(* IEC 61131-3 sources: STAR-PLC-Agent/results/raw/four_group_20261114/star_deepseek_v4/PUB020/generation/sim_00, 1 file *)

(* ---- test_program.st ---- *)
PROGRAM PLC_PRG
VAR
 BenchStep : UDINT := 0;
 BenchCalls : UDINT := 0;
 BenchDone : BOOL := FALSE;
 BenchUut0 : FB_Task;
 BenchUut1 : FB_Task;
 TraceIn_Mode : ARRAY[0..14] OF BOOL;
 TraceIn_ForwardButton : ARRAY[0..14] OF BOOL;
 TraceIn_ReverseButton : ARRAY[0..14] OF BOOL;
 TraceIn_SensorFeed : ARRAY[0..14] OF BOOL;
 TraceIn_SensorWash : ARRAY[0..14] OF BOOL;
 TraceIn_SensorWeight : ARRAY[0..14] OF BOOL;
 TraceIn_SensorFiring : ARRAY[0..14] OF BOOL;
 TraceIn_SensorOutput : ARRAY[0..14] OF BOOL;
 TraceIn_washComplete : ARRAY[0..14] OF BOOL;
 TraceIn_weightComplete : ARRAY[0..14] OF BOOL;
 TraceIn_weight : ARRAY[0..14] OF REAL;
 TraceIn_firingComplete : ARRAY[0..14] OF BOOL;
 TraceOut_MotorForward : ARRAY[0..14] OF BOOL;
 TraceOut_MotorReverse : ARRAY[0..14] OF BOOL;
 TraceOut_kick : ARRAY[0..14] OF BOOL;
 TraceOut_CompletionLight : ARRAY[0..14] OF BOOL;
 TraceOut_firingTemp : ARRAY[0..14] OF REAL;
END_VAR

IF NOT BenchDone THEN
 CASE BenchStep OF
 0:
   BenchUut0.Mode := TRUE;
   BenchUut0.ForwardButton := FALSE;
   BenchUut0.ReverseButton := FALSE;
   BenchUut0.SensorFeed := TRUE;
   BenchUut0.SensorWash := FALSE;
   BenchUut0.SensorWeight := FALSE;
   BenchUut0.SensorFiring := FALSE;
   BenchUut0.SensorOutput := FALSE;
   BenchUut0.washComplete := FALSE;
   BenchUut0.weightComplete := FALSE;
   BenchUut0.weight := REAL#0.0;
   BenchUut0.firingComplete := FALSE;
   TraceIn_Mode[0] := BenchUut0.Mode;
   TraceIn_ForwardButton[0] := BenchUut0.ForwardButton;
   TraceIn_ReverseButton[0] := BenchUut0.ReverseButton;
   TraceIn_SensorFeed[0] := BenchUut0.SensorFeed;
   TraceIn_SensorWash[0] := BenchUut0.SensorWash;
   TraceIn_SensorWeight[0] := BenchUut0.SensorWeight;
   TraceIn_SensorFiring[0] := BenchUut0.SensorFiring;
   TraceIn_SensorOutput[0] := BenchUut0.SensorOutput;
   TraceIn_washComplete[0] := BenchUut0.washComplete;
   TraceIn_weightComplete[0] := BenchUut0.weightComplete;
   TraceIn_weight[0] := BenchUut0.weight;
   TraceIn_firingComplete[0] := BenchUut0.firingComplete;
   BenchUut0();
   TraceOut_MotorForward[0] := BenchUut0.MotorForward;
   TraceOut_MotorReverse[0] := BenchUut0.MotorReverse;
   TraceOut_kick[0] := BenchUut0.kick;
   TraceOut_CompletionLight[0] := BenchUut0.CompletionLight;
   TraceOut_firingTemp[0] := BenchUut0.firingTemp;
   BenchCalls := BenchCalls + 1;
 1:
   BenchUut0.Mode := TRUE;
   BenchUut0.ForwardButton := FALSE;
   BenchUut0.ReverseButton := FALSE;
   BenchUut0.SensorFeed := FALSE;
   BenchUut0.SensorWash := TRUE;
   BenchUut0.SensorWeight := FALSE;
   BenchUut0.SensorFiring := FALSE;
   BenchUut0.SensorOutput := FALSE;
   BenchUut0.washComplete := FALSE;
   BenchUut0.weightComplete := FALSE;
   BenchUut0.weight := REAL#0.0;
   BenchUut0.firingComplete := FALSE;
   TraceIn_Mode[1] := BenchUut0.Mode;
   TraceIn_ForwardButton[1] := BenchUut0.ForwardButton;
   TraceIn_ReverseButton[1] := BenchUut0.ReverseButton;
   TraceIn_SensorFeed[1] := BenchUut0.SensorFeed;
   TraceIn_SensorWash[1] := BenchUut0.SensorWash;
   TraceIn_SensorWeight[1] := BenchUut0.SensorWeight;
   TraceIn_SensorFiring[1] := BenchUut0.SensorFiring;
   TraceIn_SensorOutput[1] := BenchUut0.SensorOutput;
   TraceIn_washComplete[1] := BenchUut0.washComplete;
   TraceIn_weightComplete[1] := BenchUut0.weightComplete;
   TraceIn_weight[1] := BenchUut0.weight;
   TraceIn_firingComplete[1] := BenchUut0.firingComplete;
   BenchUut0();
   TraceOut_MotorForward[1] := BenchUut0.MotorForward;
   TraceOut_MotorReverse[1] := BenchUut0.MotorReverse;
   TraceOut_kick[1] := BenchUut0.kick;
   TraceOut_CompletionLight[1] := BenchUut0.CompletionLight;
   TraceOut_firingTemp[1] := BenchUut0.firingTemp;
   BenchCalls := BenchCalls + 1;
 2:
   BenchUut0.Mode := TRUE;
   BenchUut0.ForwardButton := FALSE;
   BenchUut0.ReverseButton := FALSE;
   BenchUut0.SensorFeed := FALSE;
   BenchUut0.SensorWash := TRUE;
   BenchUut0.SensorWeight := FALSE;
   BenchUut0.SensorFiring := FALSE;
   BenchUut0.SensorOutput := FALSE;
   BenchUut0.washComplete := TRUE;
   BenchUut0.weightComplete := FALSE;
   BenchUut0.weight := REAL#0.0;
   BenchUut0.firingComplete := FALSE;
   TraceIn_Mode[2] := BenchUut0.Mode;
   TraceIn_ForwardButton[2] := BenchUut0.ForwardButton;
   TraceIn_ReverseButton[2] := BenchUut0.ReverseButton;
   TraceIn_SensorFeed[2] := BenchUut0.SensorFeed;
   TraceIn_SensorWash[2] := BenchUut0.SensorWash;
   TraceIn_SensorWeight[2] := BenchUut0.SensorWeight;
   TraceIn_SensorFiring[2] := BenchUut0.SensorFiring;
   TraceIn_SensorOutput[2] := BenchUut0.SensorOutput;
   TraceIn_washComplete[2] := BenchUut0.washComplete;
   TraceIn_weightComplete[2] := BenchUut0.weightComplete;
   TraceIn_weight[2] := BenchUut0.weight;
   TraceIn_firingComplete[2] := BenchUut0.firingComplete;
   BenchUut0();
   TraceOut_MotorForward[2] := BenchUut0.MotorForward;
   TraceOut_MotorReverse[2] := BenchUut0.MotorReverse;
   TraceOut_kick[2] := BenchUut0.kick;
   TraceOut_CompletionLight[2] := BenchUut0.CompletionLight;
   TraceOut_firingTemp[2] := BenchUut0.firingTemp;
   BenchCalls := BenchCalls + 1;
 3:
   BenchUut0.Mode := TRUE;
   BenchUut0.ForwardButton := FALSE;
   BenchUut0.ReverseButton := FALSE;
   BenchUut0.SensorFeed := FALSE;
   BenchUut0.SensorWash := FALSE;
   BenchUut0.SensorWeight := TRUE;
   BenchUut0.SensorFiring := FALSE;
   BenchUut0.SensorOutput := FALSE;
   BenchUut0.washComplete := FALSE;
   BenchUut0.weightComplete := FALSE;
   BenchUut0.weight := REAL#0.0;
   BenchUut0.firingComplete := FALSE;
   TraceIn_Mode[3] := BenchUut0.Mode;
   TraceIn_ForwardButton[3] := BenchUut0.ForwardButton;
   TraceIn_ReverseButton[3] := BenchUut0.ReverseButton;
   TraceIn_SensorFeed[3] := BenchUut0.SensorFeed;
   TraceIn_SensorWash[3] := BenchUut0.SensorWash;
   TraceIn_SensorWeight[3] := BenchUut0.SensorWeight;
   TraceIn_SensorFiring[3] := BenchUut0.SensorFiring;
   TraceIn_SensorOutput[3] := BenchUut0.SensorOutput;
   TraceIn_washComplete[3] := BenchUut0.washComplete;
   TraceIn_weightComplete[3] := BenchUut0.weightComplete;
   TraceIn_weight[3] := BenchUut0.weight;
   TraceIn_firingComplete[3] := BenchUut0.firingComplete;
   BenchUut0();
   TraceOut_MotorForward[3] := BenchUut0.MotorForward;
   TraceOut_MotorReverse[3] := BenchUut0.MotorReverse;
   TraceOut_kick[3] := BenchUut0.kick;
   TraceOut_CompletionLight[3] := BenchUut0.CompletionLight;
   TraceOut_firingTemp[3] := BenchUut0.firingTemp;
   BenchCalls := BenchCalls + 1;
 4:
   BenchUut0.Mode := TRUE;
   BenchUut0.ForwardButton := FALSE;
   BenchUut0.ReverseButton := FALSE;
   BenchUut0.SensorFeed := FALSE;
   BenchUut0.SensorWash := FALSE;
   BenchUut0.SensorWeight := TRUE;
   BenchUut0.SensorFiring := FALSE;
   BenchUut0.SensorOutput := FALSE;
   BenchUut0.washComplete := FALSE;
   BenchUut0.weightComplete := TRUE;
   BenchUut0.weight := REAL#200.0;
   BenchUut0.firingComplete := FALSE;
   TraceIn_Mode[4] := BenchUut0.Mode;
   TraceIn_ForwardButton[4] := BenchUut0.ForwardButton;
   TraceIn_ReverseButton[4] := BenchUut0.ReverseButton;
   TraceIn_SensorFeed[4] := BenchUut0.SensorFeed;
   TraceIn_SensorWash[4] := BenchUut0.SensorWash;
   TraceIn_SensorWeight[4] := BenchUut0.SensorWeight;
   TraceIn_SensorFiring[4] := BenchUut0.SensorFiring;
   TraceIn_SensorOutput[4] := BenchUut0.SensorOutput;
   TraceIn_washComplete[4] := BenchUut0.washComplete;
   TraceIn_weightComplete[4] := BenchUut0.weightComplete;
   TraceIn_weight[4] := BenchUut0.weight;
   TraceIn_firingComplete[4] := BenchUut0.firingComplete;
   BenchUut0();
   TraceOut_MotorForward[4] := BenchUut0.MotorForward;
   TraceOut_MotorReverse[4] := BenchUut0.MotorReverse;
   TraceOut_kick[4] := BenchUut0.kick;
   TraceOut_CompletionLight[4] := BenchUut0.CompletionLight;
   TraceOut_firingTemp[4] := BenchUut0.firingTemp;
   BenchCalls := BenchCalls + 1;
 5:
   BenchUut0.Mode := TRUE;
   BenchUut0.ForwardButton := FALSE;
   BenchUut0.ReverseButton := FALSE;
   BenchUut0.SensorFeed := FALSE;
   BenchUut0.SensorWash := FALSE;
   BenchUut0.SensorWeight := FALSE;
   BenchUut0.SensorFiring := TRUE;
   BenchUut0.SensorOutput := FALSE;
   BenchUut0.washComplete := FALSE;
   BenchUut0.weightComplete := FALSE;
   BenchUut0.weight := REAL#200.0;
   BenchUut0.firingComplete := FALSE;
   TraceIn_Mode[5] := BenchUut0.Mode;
   TraceIn_ForwardButton[5] := BenchUut0.ForwardButton;
   TraceIn_ReverseButton[5] := BenchUut0.ReverseButton;
   TraceIn_SensorFeed[5] := BenchUut0.SensorFeed;
   TraceIn_SensorWash[5] := BenchUut0.SensorWash;
   TraceIn_SensorWeight[5] := BenchUut0.SensorWeight;
   TraceIn_SensorFiring[5] := BenchUut0.SensorFiring;
   TraceIn_SensorOutput[5] := BenchUut0.SensorOutput;
   TraceIn_washComplete[5] := BenchUut0.washComplete;
   TraceIn_weightComplete[5] := BenchUut0.weightComplete;
   TraceIn_weight[5] := BenchUut0.weight;
   TraceIn_firingComplete[5] := BenchUut0.firingComplete;
   BenchUut0();
   TraceOut_MotorForward[5] := BenchUut0.MotorForward;
   TraceOut_MotorReverse[5] := BenchUut0.MotorReverse;
   TraceOut_kick[5] := BenchUut0.kick;
   TraceOut_CompletionLight[5] := BenchUut0.CompletionLight;
   TraceOut_firingTemp[5] := BenchUut0.firingTemp;
   BenchCalls := BenchCalls + 1;
 6:
   BenchUut0.Mode := TRUE;
   BenchUut0.ForwardButton := FALSE;
   BenchUut0.ReverseButton := FALSE;
   BenchUut0.SensorFeed := FALSE;
   BenchUut0.SensorWash := FALSE;
   BenchUut0.SensorWeight := FALSE;
   BenchUut0.SensorFiring := TRUE;
   BenchUut0.SensorOutput := FALSE;
   BenchUut0.washComplete := FALSE;
   BenchUut0.weightComplete := FALSE;
   BenchUut0.weight := REAL#200.0;
   BenchUut0.firingComplete := TRUE;
   TraceIn_Mode[6] := BenchUut0.Mode;
   TraceIn_ForwardButton[6] := BenchUut0.ForwardButton;
   TraceIn_ReverseButton[6] := BenchUut0.ReverseButton;
   TraceIn_SensorFeed[6] := BenchUut0.SensorFeed;
   TraceIn_SensorWash[6] := BenchUut0.SensorWash;
   TraceIn_SensorWeight[6] := BenchUut0.SensorWeight;
   TraceIn_SensorFiring[6] := BenchUut0.SensorFiring;
   TraceIn_SensorOutput[6] := BenchUut0.SensorOutput;
   TraceIn_washComplete[6] := BenchUut0.washComplete;
   TraceIn_weightComplete[6] := BenchUut0.weightComplete;
   TraceIn_weight[6] := BenchUut0.weight;
   TraceIn_firingComplete[6] := BenchUut0.firingComplete;
   BenchUut0();
   TraceOut_MotorForward[6] := BenchUut0.MotorForward;
   TraceOut_MotorReverse[6] := BenchUut0.MotorReverse;
   TraceOut_kick[6] := BenchUut0.kick;
   TraceOut_CompletionLight[6] := BenchUut0.CompletionLight;
   TraceOut_firingTemp[6] := BenchUut0.firingTemp;
   BenchCalls := BenchCalls + 1;
 7:
   BenchUut0.Mode := TRUE;
   BenchUut0.ForwardButton := FALSE;
   BenchUut0.ReverseButton := FALSE;
   BenchUut0.SensorFeed := FALSE;
   BenchUut0.SensorWash := FALSE;
   BenchUut0.SensorWeight := FALSE;
   BenchUut0.SensorFiring := FALSE;
   BenchUut0.SensorOutput := TRUE;
   BenchUut0.washComplete := FALSE;
   BenchUut0.weightComplete := FALSE;
   BenchUut0.weight := REAL#200.0;
   BenchUut0.firingComplete := FALSE;
   TraceIn_Mode[7] := BenchUut0.Mode;
   TraceIn_ForwardButton[7] := BenchUut0.ForwardButton;
   TraceIn_ReverseButton[7] := BenchUut0.ReverseButton;
   TraceIn_SensorFeed[7] := BenchUut0.SensorFeed;
   TraceIn_SensorWash[7] := BenchUut0.SensorWash;
   TraceIn_SensorWeight[7] := BenchUut0.SensorWeight;
   TraceIn_SensorFiring[7] := BenchUut0.SensorFiring;
   TraceIn_SensorOutput[7] := BenchUut0.SensorOutput;
   TraceIn_washComplete[7] := BenchUut0.washComplete;
   TraceIn_weightComplete[7] := BenchUut0.weightComplete;
   TraceIn_weight[7] := BenchUut0.weight;
   TraceIn_firingComplete[7] := BenchUut0.firingComplete;
   BenchUut0();
   TraceOut_MotorForward[7] := BenchUut0.MotorForward;
   TraceOut_MotorReverse[7] := BenchUut0.MotorReverse;
   TraceOut_kick[7] := BenchUut0.kick;
   TraceOut_CompletionLight[7] := BenchUut0.CompletionLight;
   TraceOut_firingTemp[7] := BenchUut0.firingTemp;
   BenchCalls := BenchCalls + 1;
 8:
   BenchUut1.Mode := TRUE;
   BenchUut1.ForwardButton := FALSE;
   BenchUut1.ReverseButton := FALSE;
   BenchUut1.SensorFeed := TRUE;
   BenchUut1.SensorWash := FALSE;
   BenchUut1.SensorWeight := FALSE;
   BenchUut1.SensorFiring := FALSE;
   BenchUut1.SensorOutput := FALSE;
   BenchUut1.washComplete := FALSE;
   BenchUut1.weightComplete := FALSE;
   BenchUut1.weight := REAL#0.0;
   BenchUut1.firingComplete := FALSE;
   TraceIn_Mode[8] := BenchUut1.Mode;
   TraceIn_ForwardButton[8] := BenchUut1.ForwardButton;
   TraceIn_ReverseButton[8] := BenchUut1.ReverseButton;
   TraceIn_SensorFeed[8] := BenchUut1.SensorFeed;
   TraceIn_SensorWash[8] := BenchUut1.SensorWash;
   TraceIn_SensorWeight[8] := BenchUut1.SensorWeight;
   TraceIn_SensorFiring[8] := BenchUut1.SensorFiring;
   TraceIn_SensorOutput[8] := BenchUut1.SensorOutput;
   TraceIn_washComplete[8] := BenchUut1.washComplete;
   TraceIn_weightComplete[8] := BenchUut1.weightComplete;
   TraceIn_weight[8] := BenchUut1.weight;
   TraceIn_firingComplete[8] := BenchUut1.firingComplete;
   BenchUut1();
   TraceOut_MotorForward[8] := BenchUut1.MotorForward;
   TraceOut_MotorReverse[8] := BenchUut1.MotorReverse;
   TraceOut_kick[8] := BenchUut1.kick;
   TraceOut_CompletionLight[8] := BenchUut1.CompletionLight;
   TraceOut_firingTemp[8] := BenchUut1.firingTemp;
   BenchCalls := BenchCalls + 1;
 9:
   BenchUut1.Mode := TRUE;
   BenchUut1.ForwardButton := FALSE;
   BenchUut1.ReverseButton := FALSE;
   BenchUut1.SensorFeed := FALSE;
   BenchUut1.SensorWash := TRUE;
   BenchUut1.SensorWeight := FALSE;
   BenchUut1.SensorFiring := FALSE;
   BenchUut1.SensorOutput := FALSE;
   BenchUut1.washComplete := FALSE;
   BenchUut1.weightComplete := FALSE;
   BenchUut1.weight := REAL#0.0;
   BenchUut1.firingComplete := FALSE;
   TraceIn_Mode[9] := BenchUut1.Mode;
   TraceIn_ForwardButton[9] := BenchUut1.ForwardButton;
   TraceIn_ReverseButton[9] := BenchUut1.ReverseButton;
   TraceIn_SensorFeed[9] := BenchUut1.SensorFeed;
   TraceIn_SensorWash[9] := BenchUut1.SensorWash;
   TraceIn_SensorWeight[9] := BenchUut1.SensorWeight;
   TraceIn_SensorFiring[9] := BenchUut1.SensorFiring;
   TraceIn_SensorOutput[9] := BenchUut1.SensorOutput;
   TraceIn_washComplete[9] := BenchUut1.washComplete;
   TraceIn_weightComplete[9] := BenchUut1.weightComplete;
   TraceIn_weight[9] := BenchUut1.weight;
   TraceIn_firingComplete[9] := BenchUut1.firingComplete;
   BenchUut1();
   TraceOut_MotorForward[9] := BenchUut1.MotorForward;
   TraceOut_MotorReverse[9] := BenchUut1.MotorReverse;
   TraceOut_kick[9] := BenchUut1.kick;
   TraceOut_CompletionLight[9] := BenchUut1.CompletionLight;
   TraceOut_firingTemp[9] := BenchUut1.firingTemp;
   BenchCalls := BenchCalls + 1;
 10:
   BenchUut1.Mode := TRUE;
   BenchUut1.ForwardButton := FALSE;
   BenchUut1.ReverseButton := FALSE;
   BenchUut1.SensorFeed := FALSE;
   BenchUut1.SensorWash := TRUE;
   BenchUut1.SensorWeight := FALSE;
   BenchUut1.SensorFiring := FALSE;
   BenchUut1.SensorOutput := FALSE;
   BenchUut1.washComplete := TRUE;
   BenchUut1.weightComplete := FALSE;
   BenchUut1.weight := REAL#0.0;
   BenchUut1.firingComplete := FALSE;
   TraceIn_Mode[10] := BenchUut1.Mode;
   TraceIn_ForwardButton[10] := BenchUut1.ForwardButton;
   TraceIn_ReverseButton[10] := BenchUut1.ReverseButton;
   TraceIn_SensorFeed[10] := BenchUut1.SensorFeed;
   TraceIn_SensorWash[10] := BenchUut1.SensorWash;
   TraceIn_SensorWeight[10] := BenchUut1.SensorWeight;
   TraceIn_SensorFiring[10] := BenchUut1.SensorFiring;
   TraceIn_SensorOutput[10] := BenchUut1.SensorOutput;
   TraceIn_washComplete[10] := BenchUut1.washComplete;
   TraceIn_weightComplete[10] := BenchUut1.weightComplete;
   TraceIn_weight[10] := BenchUut1.weight;
   TraceIn_firingComplete[10] := BenchUut1.firingComplete;
   BenchUut1();
   TraceOut_MotorForward[10] := BenchUut1.MotorForward;
   TraceOut_MotorReverse[10] := BenchUut1.MotorReverse;
   TraceOut_kick[10] := BenchUut1.kick;
   TraceOut_CompletionLight[10] := BenchUut1.CompletionLight;
   TraceOut_firingTemp[10] := BenchUut1.firingTemp;
   BenchCalls := BenchCalls + 1;
 11:
   BenchUut1.Mode := TRUE;
   BenchUut1.ForwardButton := FALSE;
   BenchUut1.ReverseButton := FALSE;
   BenchUut1.SensorFeed := FALSE;
   BenchUut1.SensorWash := FALSE;
   BenchUut1.SensorWeight := TRUE;
   BenchUut1.SensorFiring := FALSE;
   BenchUut1.SensorOutput := FALSE;
   BenchUut1.washComplete := FALSE;
   BenchUut1.weightComplete := FALSE;
   BenchUut1.weight := REAL#0.0;
   BenchUut1.firingComplete := FALSE;
   TraceIn_Mode[11] := BenchUut1.Mode;
   TraceIn_ForwardButton[11] := BenchUut1.ForwardButton;
   TraceIn_ReverseButton[11] := BenchUut1.ReverseButton;
   TraceIn_SensorFeed[11] := BenchUut1.SensorFeed;
   TraceIn_SensorWash[11] := BenchUut1.SensorWash;
   TraceIn_SensorWeight[11] := BenchUut1.SensorWeight;
   TraceIn_SensorFiring[11] := BenchUut1.SensorFiring;
   TraceIn_SensorOutput[11] := BenchUut1.SensorOutput;
   TraceIn_washComplete[11] := BenchUut1.washComplete;
   TraceIn_weightComplete[11] := BenchUut1.weightComplete;
   TraceIn_weight[11] := BenchUut1.weight;
   TraceIn_firingComplete[11] := BenchUut1.firingComplete;
   BenchUut1();
   TraceOut_MotorForward[11] := BenchUut1.MotorForward;
   TraceOut_MotorReverse[11] := BenchUut1.MotorReverse;
   TraceOut_kick[11] := BenchUut1.kick;
   TraceOut_CompletionLight[11] := BenchUut1.CompletionLight;
   TraceOut_firingTemp[11] := BenchUut1.firingTemp;
   BenchCalls := BenchCalls + 1;
 12:
   BenchUut1.Mode := TRUE;
   BenchUut1.ForwardButton := FALSE;
   BenchUut1.ReverseButton := FALSE;
   BenchUut1.SensorFeed := FALSE;
   BenchUut1.SensorWash := FALSE;
   BenchUut1.SensorWeight := TRUE;
   BenchUut1.SensorFiring := FALSE;
   BenchUut1.SensorOutput := FALSE;
   BenchUut1.washComplete := FALSE;
   BenchUut1.weightComplete := TRUE;
   BenchUut1.weight := REAL#200.1;
   BenchUut1.firingComplete := FALSE;
   TraceIn_Mode[12] := BenchUut1.Mode;
   TraceIn_ForwardButton[12] := BenchUut1.ForwardButton;
   TraceIn_ReverseButton[12] := BenchUut1.ReverseButton;
   TraceIn_SensorFeed[12] := BenchUut1.SensorFeed;
   TraceIn_SensorWash[12] := BenchUut1.SensorWash;
   TraceIn_SensorWeight[12] := BenchUut1.SensorWeight;
   TraceIn_SensorFiring[12] := BenchUut1.SensorFiring;
   TraceIn_SensorOutput[12] := BenchUut1.SensorOutput;
   TraceIn_washComplete[12] := BenchUut1.washComplete;
   TraceIn_weightComplete[12] := BenchUut1.weightComplete;
   TraceIn_weight[12] := BenchUut1.weight;
   TraceIn_firingComplete[12] := BenchUut1.firingComplete;
   BenchUut1();
   TraceOut_MotorForward[12] := BenchUut1.MotorForward;
   TraceOut_MotorReverse[12] := BenchUut1.MotorReverse;
   TraceOut_kick[12] := BenchUut1.kick;
   TraceOut_CompletionLight[12] := BenchUut1.CompletionLight;
   TraceOut_firingTemp[12] := BenchUut1.firingTemp;
   BenchCalls := BenchCalls + 1;
 13:
   BenchUut1.Mode := TRUE;
   BenchUut1.ForwardButton := FALSE;
   BenchUut1.ReverseButton := FALSE;
   BenchUut1.SensorFeed := FALSE;
   BenchUut1.SensorWash := FALSE;
   BenchUut1.SensorWeight := FALSE;
   BenchUut1.SensorFiring := FALSE;
   BenchUut1.SensorOutput := FALSE;
   BenchUut1.washComplete := FALSE;
   BenchUut1.weightComplete := FALSE;
   BenchUut1.weight := REAL#200.1;
   BenchUut1.firingComplete := FALSE;
   TraceIn_Mode[13] := BenchUut1.Mode;
   TraceIn_ForwardButton[13] := BenchUut1.ForwardButton;
   TraceIn_ReverseButton[13] := BenchUut1.ReverseButton;
   TraceIn_SensorFeed[13] := BenchUut1.SensorFeed;
   TraceIn_SensorWash[13] := BenchUut1.SensorWash;
   TraceIn_SensorWeight[13] := BenchUut1.SensorWeight;
   TraceIn_SensorFiring[13] := BenchUut1.SensorFiring;
   TraceIn_SensorOutput[13] := BenchUut1.SensorOutput;
   TraceIn_washComplete[13] := BenchUut1.washComplete;
   TraceIn_weightComplete[13] := BenchUut1.weightComplete;
   TraceIn_weight[13] := BenchUut1.weight;
   TraceIn_firingComplete[13] := BenchUut1.firingComplete;
   BenchUut1();
   TraceOut_MotorForward[13] := BenchUut1.MotorForward;
   TraceOut_MotorReverse[13] := BenchUut1.MotorReverse;
   TraceOut_kick[13] := BenchUut1.kick;
   TraceOut_CompletionLight[13] := BenchUut1.CompletionLight;
   TraceOut_firingTemp[13] := BenchUut1.firingTemp;
   BenchCalls := BenchCalls + 1;
 14:
   BenchUut1.Mode := TRUE;
   BenchUut1.ForwardButton := FALSE;
   BenchUut1.ReverseButton := FALSE;
   BenchUut1.SensorFeed := TRUE;
   BenchUut1.SensorWash := FALSE;
   BenchUut1.SensorWeight := FALSE;
   BenchUut1.SensorFiring := FALSE;
   BenchUut1.SensorOutput := FALSE;
   BenchUut1.washComplete := FALSE;
   BenchUut1.weightComplete := FALSE;
   BenchUut1.weight := REAL#0.0;
   BenchUut1.firingComplete := FALSE;
   TraceIn_Mode[14] := BenchUut1.Mode;
   TraceIn_ForwardButton[14] := BenchUut1.ForwardButton;
   TraceIn_ReverseButton[14] := BenchUut1.ReverseButton;
   TraceIn_SensorFeed[14] := BenchUut1.SensorFeed;
   TraceIn_SensorWash[14] := BenchUut1.SensorWash;
   TraceIn_SensorWeight[14] := BenchUut1.SensorWeight;
   TraceIn_SensorFiring[14] := BenchUut1.SensorFiring;
   TraceIn_SensorOutput[14] := BenchUut1.SensorOutput;
   TraceIn_washComplete[14] := BenchUut1.washComplete;
   TraceIn_weightComplete[14] := BenchUut1.weightComplete;
   TraceIn_weight[14] := BenchUut1.weight;
   TraceIn_firingComplete[14] := BenchUut1.firingComplete;
   BenchUut1();
   TraceOut_MotorForward[14] := BenchUut1.MotorForward;
   TraceOut_MotorReverse[14] := BenchUut1.MotorReverse;
   TraceOut_kick[14] := BenchUut1.kick;
   TraceOut_CompletionLight[14] := BenchUut1.CompletionLight;
   TraceOut_firingTemp[14] := BenchUut1.firingTemp;
   BenchCalls := BenchCalls + 1;
 END_CASE;
 BenchStep := BenchStep + 1;
 IF BenchStep >= 15 THEN BenchDone := TRUE; END_IF;
END_IF;
END_PROGRAM
